FUNCTION F_STRING_TO_BYTES_TERM (* STRING mit Textende 16#00 in ein BYTE-Array kopieren (z. B. fuer AlPgnTxNew_TP), Rest 16#FF *)
  (* Standard: 61499-1; Description: Copyright (c) 2026 HR Agrartechnik GmbH This program and the accompanying materials are made available under the terms of the Eclipse Public License 2.0 which is available at https://www.eclipse.org/legal/epl-2.0/ SPDX-License-Identifier: EPL-2.0 *)
  (* Version 1.0, 2026-11-26, Franz Höpfinger, HR Agrartechnik GmbH, Initial Version - wie F_STRING_TO_BYTES 1.1 *)
  PACKAGE logiBUS::utils::dyn_arr;
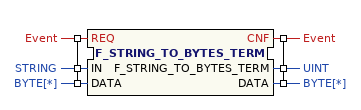
  EVENT_INPUT
    REQ WITH IN, DATA;
  END_EVENT
  EVENT_OUTPUT
    CNF WITH F_STRING_TO_BYTES_TERM, DATA;
  END_EVENT
  VAR_INPUT
    IN : STRING; (* Text, je Zeichen 1 Byte *)
  END_VAR
  VAR_OUTPUT
    F_STRING_TO_BYTES_TERM : UINT; (* Zeichen + 16#00, hoechstens die Groesse von DATA *)
  END_VAR
  VAR_IN_OUT
    DATA : ARRAY [*] OF BYTE; (* Zielpuffer, z. B. von PROVIDE_ARR_xxxx_BYTE, wird ganz beschrieben *)
  END_VAR
  BODY IN ST:
PACKAGE logiBUS::utils::dyn_arr;

(* STRING in ein BYTE-Array kopieren: Zeichen, dann 16#00 (falls Platz), Rest 16#FF *)
FUNCTION F_STRING_TO_BYTES_TERM : UINT

VAR_INPUT
	IN : STRING; // Text, je Zeichen 1 Byte
END_VAR

VAR_IN_OUT
	DATA : ARRAY[*] OF BYTE; // Zielpuffer
END_VAR

VAR_TEMP
	lo : DINT; // erster Index von DATA
	cap : DINT; // Groesse von DATA
	n : DINT; // Anzahl zu kopierender Zeichen
	i : DINT; // Laufindex
END_VAR

lo := LOWER_BOUND(DATA, 1);
cap := UPPER_BOUND(DATA, 1) - lo + 1;
n := LEN(IN);
IF n < 0 THEN
	n := 0;
END_IF;
IF n > cap THEN
	n := cap;
END_IF;
FOR i := 1 TO cap DO
	DATA[lo + i - 1] := BYTE#16#FF; // nicht genutzte Bytes wie bei J1939/ISOBUS ueblich
END_FOR;
FOR i := 1 TO n DO
	DATA[lo + i - 1] := CHAR_TO_BYTE(IN[i]);
END_FOR;
IF n < cap THEN
	DATA[lo + n] := BYTE#16#00; // Textende
	n := n + 1;
END_IF;
F_STRING_TO_BYTES_TERM := DINT_TO_UINT(n);

END_FUNCTION
  END_BODY
END_FUNCTION
